// TIA Portal V21 export
// export: Created 2026-08-21T20:18:52.6792221Z, ExportSetting None, DisplayName Totally Integrated Automation Portal, DisplayVersion V21, DisplayName STEP 7 Professional, DisplayVersion V21, DisplayName STEP 7 Safety, DisplayVersion V21, DisplayName Tech WebApplication, DisplayVersion V21, DisplayName WinCC Basic/Comfort/Advanced, DisplayVersion V21, DisplayName WinCC Professional, DisplayVersion V21, DisplayName WinCC Unified, DisplayVersion V21
FUNCTION_BLOCK "ServiceMediumParameterHMI"   // FB1754, SCL
TITLE = ServiceMediumParameterHMI
{ S7_Optimized_Access := 'TRUE' }
AUTHOR : Siemens AG
FAMILY : ServiceControl
VERSION : 4.0
// { "TagName" : "" , "TagDescription" : "" }
// stored: MemoryReserve 100, SetENOAutomatically false
   VAR_INPUT
      Id { ExternalAccessible := 'False'; ExternalVisible := 'False'; ExternalWritable := 'False'} : USInt;   // Service parameter ID
      Setup { ExternalAccessible := 'False'; ExternalVisible := 'False'; ExternalWritable := 'False'} : DB_ANY;   // Setup DB used for the service
      ProcedureCur { ExternalAccessible := 'False'; ExternalVisible := 'False'; ExternalWritable := 'False'} : DWord;   // Current Procedure Number
      ProcedureReq { ExternalAccessible := 'False'; ExternalVisible := 'False'; ExternalWritable := 'False'} : DWord;   // Required Procedure Numbar
   END_VAR
   VAR_IN_OUT
      ConfigurationParameterAnalog : Array[*] of "UDT_MTP_AnaServParam";   // Analog configuration parameter
      ConfigurationParameterDigital : Array[*] of "UDT_MTP_DIntServParam";   // Digital configuration parameter
      ConfigurationParameterBinary : Array[*] of "UDT_MTP_BinServParam";   // Binary configuration parameter
      ConfigurationParameterString : Array[*] of "UDT_MTP_StringServParam";   // String configuration parameter
      ProcedureParameterAnalog : Array[*] of "UDT_MTP_AnaServParam";   // Analog configuration parameter / Analog procedure parameter
      ProcedureParameterDigital : Array[*] of "UDT_MTP_DIntServParam";   // Digital configuration parameter / Digital procedure parameter
      ProcedureParameterBinary : Array[*] of "UDT_MTP_BinServParam";   // Binary configuration parameter / Binary procedure parameter
      ProcedureParameterString : Array[*] of "UDT_MTP_StringServParam";   // String configuration parameter / String procedure parameter
      ProcessValueInAnalog : Array[*] of "UDT_MTP_AnaProcessValueIn";   // Analog process value in
      ProcessValueInDigital : Array[*] of "UDT_MTP_DIntProcessValueIn";   // Digital process value in
      ProcessValueInBinary : Array[*] of "UDT_MTP_BinProcessValueIn";   // Binary process value in
      ProcessValueInString : Array[*] of "UDT_MTP_StringProcessValueIn";   // String process value in
      ProcessValueOutAnalog : Array[*] of "UDT_MTP_AnaProcessValueOut";   // Analog process value out
      ProcessValueOutDigital : Array[*] of "UDT_MTP_DIntProcessValueOut";   // Digital process value out
      ProcessValueOutBinary : Array[*] of "UDT_MTP_BinProcessValueOut";   // Binary process value out
      ProcessValueOutString : Array[*] of "UDT_MTP_StringProcessValueOut";   // String process value out
      ReportValueAnalog : Array[*] of "UDT_MTP_AnaReportValue";   // Analog report value
      ReportValueDigital : Array[*] of "UDT_MTP_DIntReportValue";   // Digital report value
      ReportValueBinary : Array[*] of "UDT_MTP_BinReportValue";   // Binary report value
      ReportValueString : Array[*] of "UDT_MTP_StringReportValue";   // String report value
   END_VAR
   VAR
      statTotalConfigParameters { ExternalAccessible := 'False'; ExternalVisible := 'False'; ExternalWritable := 'False'} : Int;   // Total used configuration parameter
      statTotalProcedureParameters { ExternalAccessible := 'False'; ExternalVisible := 'False'; ExternalWritable := 'False'} : Int;   // Total used procedure parameter
      statTotalProcessInValues { ExternalAccessible := 'False'; ExternalVisible := 'False'; ExternalWritable := 'False'} : Int;   // Total used process in values
      statTotalProcessOutValues { ExternalAccessible := 'False'; ExternalVisible := 'False'; ExternalWritable := 'False'} : Int;   // Total used process Out values
      statTotalReportValues { ExternalAccessible := 'False'; ExternalVisible := 'False'; ExternalWritable := 'False'} : Int;   // Total used Report values
      StatConfigAnalog { ExternalAccessible := 'False'; ExternalVisible := 'False'; ExternalWritable := 'False'} : Array[0..#MAPPED_CONFIG_ANALOG] of "UDT_Service_AnaServParam";   // Writable Config analog parameters
      StatConfigDigital { ExternalAccessible := 'False'; ExternalVisible := 'False'; ExternalWritable := 'False'} : Array[0..#MAPPED_CONFIG_DIGITAL] of "UDT_Service_DintServParam";   // Writable Config digital parameters
      StatConfigBinary { ExternalAccessible := 'False'; ExternalVisible := 'False'; ExternalWritable := 'False'} : Array[0..#MAPPED_CONFIG_BINARY] of "UDT_Service_BinServParam";   // Writable Config binary parameters
      StatConfigString { ExternalAccessible := 'False'; ExternalVisible := 'False'; ExternalWritable := 'False'} : Array[0..#MAPPED_CONFIG_STRING] of "UDT_Service_StringServParam";   // Writable Config string parameters
      StatProcedureAnalog { ExternalAccessible := 'False'; ExternalVisible := 'False'; ExternalWritable := 'False'} : Array[0..#MAPPED_PROCEDURE_ANALOG] of "UDT_Service_AnaServParam";   // Writable Config analog parameters
      StatProcedureDigital { ExternalAccessible := 'False'; ExternalVisible := 'False'; ExternalWritable := 'False'} : Array[0..#MAPPED_PROCEDURE_DIGITAL] of "UDT_Service_DintServParam";   // Writable Config digital parameters
      StatProcedureBinary { ExternalAccessible := 'False'; ExternalVisible := 'False'; ExternalWritable := 'False'} : Array[0..#MAPPED_PROCEDURE_BINARY] of "UDT_Service_BinServParam";   // Writable Config binary parameters
      StatProcedureString { ExternalAccessible := 'False'; ExternalVisible := 'False'; ExternalWritable := 'False'} : Array[0..#MAPPED_PROCEDURE_STRING] of "UDT_Service_StringServParam";   // Writable Config string parameters
      stat16ProceReqIndex { ExternalAccessible := 'False'; ExternalVisible := 'False'; ExternalWritable := 'False'} : Int;   // Requested/Prepared procedure index number
      stat16ProceCurIndex { ExternalAccessible := 'False'; ExternalVisible := 'False'; ExternalWritable := 'False'} : Int;   // current/Running procedure index number
      stat16ProcParaStartIndex { ExternalAccessible := 'False'; ExternalVisible := 'False'; ExternalWritable := 'False'} : Int;   // Procedure parameter start index value
      stat16ProcParaEndIndex { ExternalAccessible := 'False'; ExternalVisible := 'False'; ExternalWritable := 'False'} : Int;   // Procedure parameter end index value
      stat32PrecedureProcessOutMap { ExternalAccessible := 'False'; ExternalVisible := 'False'; ExternalWritable := 'False'} : DWord;   // Procedure assignment information for ProcessOut values
      stat32PrecedureProcessInMap { ExternalAccessible := 'False'; ExternalVisible := 'False'; ExternalWritable := 'False'} : DWord;   // Procedure assignment information for ProcessIn values
      stat32PrecedureReportMap { ExternalAccessible := 'False'; ExternalVisible := 'False'; ExternalWritable := 'False'} : DWord;   // Procedure assignment information for Report values
      ConfigParaType : "UDT_Service_ConfigParaIndexType";   // Index information for the configuration parameter
      ProcedureParaType : "UDT_Service_ProceParaValueIndexType";   // Index information for the procedure parameter
      ProcessInValueType : "UDT_Service_ProceParaValueIndexType";   // Index information for the process in values
      ProcessOutValueType : "UDT_Service_ProceParaValueIndexType";   // Index information for the process out values
      ReportValueType : "UDT_Service_ProceParaValueIndexType";   // Index information for the report values
      ConfigAna : Array[0..#MAPPED_CONFIG_ANALOG] of "UDT_MTP_AnaServParam";   // Configuration analog parameter
      ConfigDint : Array[0..#MAPPED_CONFIG_DIGITAL] of "UDT_MTP_DIntServParam";   // Configuration digital parameter
      ConfigBin : Array[0..#MAPPED_CONFIG_BINARY] of "UDT_MTP_BinServParam";   // Configuration binary parameter
      ConfigString : Array[0..#MAPPED_CONFIG_STRING] of "UDT_MTP_StringServParam";   // Configuration string parameter
      ProcedureAna : Array[0..#MAPPED_PROCEDURE_ANALOG] of "UDT_MTP_AnaServParam";   // Procedure analog parameter
      ProcedureDint : Array[0..#MAPPED_PROCEDURE_DIGITAL] of "UDT_MTP_DIntServParam";   // Procedure digital parameter
      ProcedureBin : Array[0..#MAPPED_PROCEDURE_BINARY] of "UDT_MTP_BinServParam";   // Procedure binary parameter
      ProcedureString : Array[0..#MAPPED_PROCEDURE_STRING] of "UDT_MTP_StringServParam";   // Procedure string parameter
      ProcessInAna : Array[0..#MAPPED_PROCESS_IN_ANALOG] of "UDT_MTP_AnaProcessValueIn";   // Process In analog values
      ProcessInDint : Array[0..#MAPPED_PROCESS_IN_DIGITAL] of "UDT_MTP_DIntProcessValueIn";   // Process In digital values
      ProcessInBin : Array[0..#MAPPED_PROCESS_IN_BINARY] of "UDT_MTP_BinProcessValueIn";   // Process In binary values
      ProcessInString : Array[0..#MAPPED_PROCESS_IN_STRING] of "UDT_MTP_StringProcessValueIn";   // Process In string values
      ProcessOutAna : Array[0..#MAPPED_PROCESS_OUT_ANALOG] of "UDT_MTP_AnaProcessValueOut";   // Process Out analog values
      ProcessOutDint : Array[0..#MAPPED_PROCESS_OUT_DIGITAL] of "UDT_MTP_DIntProcessValueOut";   // Process Out digital values
      ProcessOutBin : Array[0..#MAPPED_PROCESS_OUT_BINARY] of "UDT_MTP_BinProcessValueOut";   // Process Out binary values
      ProcessOutString : Array[0..#MAPPED_PROCESS_OUT_STRING] of "UDT_MTP_StringProcessValueOut";   // Process Out string values
      ReportAna : Array[0..#MAPPED_REPORT_ANALOG] of "UDT_MTP_AnaReportValue";   // Report analog values
      ReportDint : Array[0..#MAPPED_REPORT_DIGITAL] of "UDT_MTP_DIntReportValue";   // Report digital values
      ReportBin : Array[0..#MAPPED_REPORT_BINARY] of "UDT_MTP_BinReportValue";   // Report binary values
      ReportString : Array[0..#MAPPED_REPORT_STRING] of "UDT_MTP_StringReportValue";   // Report string values
      statInternalCurProcParameter { ExternalAccessible := 'False'; ExternalVisible := 'False'; ExternalWritable := 'False'} : Array[#PROCEDURE_PARAMETER_MIN..#PROCEDURE_PARAMETER_MAX] of "UDT_Service_Parameter";   // Internal Procedure Parameter
      statLasProcedureCur { ExternalAccessible := 'False'; ExternalVisible := 'False'; ExternalWritable := 'False'} : DWord;   // Last current procedure
      statLasProcedureReq { ExternalAccessible := 'False'; ExternalVisible := 'False'; ExternalWritable := 'False'} : DWord;   // Last Prepared procedure
      statLastReqProcedSelected { ExternalAccessible := 'False'; ExternalVisible := 'False'; ExternalWritable := 'False'} : Bool;   // Last Prepared procedure
      StatLastProceselReport { ExternalAccessible := 'False'; ExternalVisible := 'False'; ExternalWritable := 'False'} : Bool;   // Last procedure page selection in Report values FP
      StatLastProceselProcessOut { ExternalAccessible := 'False'; ExternalVisible := 'False'; ExternalWritable := 'False'} : Bool;   // Last procedure page selection in ProcessOut values FP
      StatLastProceselProcessIn { ExternalAccessible := 'False'; ExternalVisible := 'False'; ExternalWritable := 'False'} : Bool;   // Last procedure page selection in ProcessIn values FP
   END_VAR
   VAR_TEMP
      temp32TempDword1 : DWord;   // Dummy for work
      temp16IndexOfDefinition : Int;   // Index of Definition array / Internal counter variable
      temp16ParameterCMAddress : Int;   // Control module address of parameter
      temp16ParameterType : Int;   // Type of Parameter
      temp16IndexMTP : Int;   // Index of MTP array / Index fo value
      temp16IndexIO : Int;   // Index of IO array / Index fo value
      tempUsed : Array[#NUMBER_OF_CONTROLMODULES_IN_DW_MIN..#NUMBER_OF_CONTROLMODULES_IN_DW] of DWord;   // Array for input value used
      temp16TempInt1 : Int;   // Dummy for work
      temp16TempInt2 : Int;   // Dummy for work
      temp16i : Int;   // Internal counter variable
      temp16Index : Int;   // Index of value / Index fo value
      tempVariant : Variant;   // Internal work variable of type Variant
      temp16ReturnValue : Int;   // Internal work variable for Return Value
      tempSetup : "UDT_Service_ControlBlockMedium";   // Content of DB "ServiceControlBlockMediumSetup"
      tempProcStartIndex : Int;   // Procedure start index
      tempProcEndIndex : Int;   // Procedure end index
      temp16InitIndex : Int;   // Variable is used to initialize the Digital & String para index
      tempProcStartingStartIndex : Int;   // Procedure start index for Starting state
      tempProcStartingEndIndex : Int;   // Procedure end index for Starting state
      tempProcRunningStartIndex : Int;   // Procedure start index for Running state
      tempProcRunningEndIndex : Int;   // Procedure end index for Running state
      tempProcHoldingStartIndex : Int;   // Procedure start index for Holding state
      tempProcHoldingEndIndex : Int;   // Procedure end index for Holding state
      tempProcUnHoldingStartIndex : Int;   // Procedure start index for UnHolding state
      tempProcUnHoldingEndIndex : Int;   // Procedure end index for UnHolding state
      tempProcUnPausingStartIndex : Int;   // Procedure start index for Pausing state
      tempProcUnPausingEndIndex : Int;   // Procedure end index for Pausing state
      tempProcResumingStartIndex : Int;   // Procedure start index for Resuming state
      tempProcResumingEndIndex : Int;   // Procedure end index for Resuming state
      tempProcCompletingStartIndex : Int;   // Procedure start index for Completing state
      tempProcCompletingEndIndex : Int;   // Procedure end index for Completing state
      tempProcStoppingStartIndex : Int;   // Procedure start index for Stopping state
      tempProcStoppingEndIndex : Int;   // Procedure end index for Stopping state
      tempProcAbortingStartIndex : Int;   // Procedure start index for Aborting state
      tempProcAbortingEndIndex : Int;   // Procedure end index for Aborting state
      tempProcResettingStartIndex : Int;   // Procedure start index for Resetting state
      tempProcResettingEndIndex : Int;   // Procedure end index for Resetting state
      temp16IndexOfDefinitionProcessOut : Int;   // Index of Definition array / Internal counter variable
      temp16IndexOfDefinitionProcessIn : Int;   // Index of Definition array / Internal counter variable
      temp16IndexOfDefinitionReport : Int;   // Index of Definition array / Internal counter variable
      temp16IndexAnalog : Int;   // Pointer for the used analog parameter
      temp16IndexDigital : Int;   // Pointer for the used digital parameter
      temp16IndexBinary : Int;   // Pointer for the used binary parameter
      temp16IndexString : Int;   // Pointer for the used string parameter
      temp16ReturnValueOBNum : Int;   // Internal work variable for Return Value
      tempTopSi : SI_none;   // Start-up information of current OB
      tempStartSi : SI_none;   // Start-up information of last started OB
      temp16ObNo : UInt;   // OB number
      xOB_Start : Bool;   // block is running in start OB
      temp16ReturnStatus : Word;   // Internal work variable for Return Value
      tempDTLCurrentTime : DTL;   // Current time stamp
   END_VAR
   VAR CONSTANT
      CONFIG_PARAMETER_MIN : Int := 0;   // Minimum number of configuration parameters (planned number -1 due to ArrayAddressing)
      CONFIG_PARAMETER_MAX : Int := 31;   // Maximum number of configuration parameters (planned number -1 due to ArrayAddressing)
      CONFIG_PARAMETER_ANALOG_MAX : Int := 31;   // Maximum number of analog configuration parameters (planned number -1 due to ArrayAddressing)
      CONFIG_PARAMETER_DIGITAL_MAX : Int := 7;   // Maximum number of digital configuration parameters (planned number -1 due to ArrayAddressing)
      CONFIG_PARAMETER_BINARY_MAX : Int := 31;   // Maximum number of binary configuration parameters (planned number -1 due to ArrayAddressing)
      CONFIG_PARAMETER_STRING_MAX : Int := 7;   // Maximum number of string configuration parameters (planned number -1 due to ArrayAddressing)
      PROCEDURE_PARAMETER_MIN : Int := 0;   // Minimum number of procedure parameters (planned number -1 due to ArrayAddressing)
      PROCEDURE_PARAMETER_MAX : Int := 31;   // Maximum number of procedure parameters (planned number -1 due to ArrayAddressing)
      PROCEDURE_PARAMETER_ANALOG_MAX : Int := 31;   // Maximum number of analog procedure parameters (planned number -1 due to ArrayAddressing)
      PROCEDURE_PARAMETER_DIGITAL_MAX : Int := 7;   // Maximum number of digital procedure parameters (planned number -1 due to ArrayAddressing)
      PROCEDURE_PARAMETER_BINARY_MAX : Int := 31;   // Maximum number of binary procedure parameters (planned number -1 due to ArrayAddressing)
      PROCEDURE_PARAMETER_STRING_MAX : Int := 7;   // Maximum number of string procedure parameters (planned number -1 due to ArrayAddressing)
      NUMBER_OF_CONTROLMODULES_IN_DW_MIN : Int := 0;   // Number of control modules coded in DWords (planned number -1 due to ArrayAddressing)
      NUMBER_OF_CONTROLMODULES_IN_DW : Int := 0;   // Number of control modules coded in DWords (planned number -1 due to ArrayAddressing)
      NUMBER_OF_CONTROLMODULES_MIN : Int := 0;   // Number of control modules (planned number -1 due to ArrayAddressing)
      NUMBER_OF_CONTROLMODULES : Int := 29;   // Number of control modules (planned number -1 due to ArrayAddressing)
      TYPE_NONE : USInt := 0;   // No parameter
      TYPE_ANALOG : USInt := 1;   // Parameter / value type analog
      TYPE_DIGITAL : USInt := 2;   // Parameter / value type digital
      TYPE_BINARY : USInt := 3;   // Parameter / value type binary
      TYPE_STRING : USInt := 4;   // Parameter type string
      NUMBER_OF_PROCEDURES_MIN : Int := 0;   // Number of operations (planned number -1 due to ArrayAddressing)
      NUMBER_OF_PROCEDURES : Int := 15;   // Number of operations (planned number -1 due to ArrayAddressing)
      PARAMETERINDEX_MIN : Int := 0;   // Minimum number of configuration parameters (planned number -1 due to ArrayAddressing)
      PARAMETERINDEX_MAX : Int := 511;   // Maximum number of configuration parameters (planned number -1 due to ArrayAddressing)
      REPORT_VALUES_MIN : Int := 0;   // Minimum number of report values (planned number -1 due to ArrayAddressing)
      REPORT_VALUES_MAX : Int := 31;   // Maximum number of report values (planned number -1 due to ArrayAddressing)
      REPORT_VALUES_ANALOG_MAX : Int := 31;   // Maximum number of analog report values (planned number -1 due to ArrayAddressing)
      REPORT_VALUES_DIGITAL_MAX : Int := 7;   // Maximum number of digital report values (planned number -1 due to ArrayAddressing)
      REPORT_VALUES_BINARY_MAX : Int := 31;   // Maximum number of binary report values (planned number -1 due to ArrayAddressing)
      REPORT_VALUES_STRING_MAX : Int := 7;   // Maximum number of string report values (planned number -1 due to ArrayAddressing)
      PROCESS_VALUES_IN_MIN : Int := 0;   // Minimum number of process values in (planned number -1 due to ArrayAddressing)
      PROCESS_VALUES_IN_MAX : Int := 31;   // Maximum number of process values in (planned number -1 due to ArrayAddressing)
      PROCESS_VALUES_IN_ANALOG_MAX : Int := 31;   // Maximum number of analog process values in (planned number -1 due to ArrayAddressing)
      PROCESS_VALUES_IN_DIGITAL_MAX : Int := 7;   // Maximum number of digital process values in (planned number -1 due to ArrayAddressing)
      PROCESS_VALUES_IN_BINARY_MAX : Int := 31;   // Maximum number of binary process values in (planned number -1 due to ArrayAddressing)
      PROCESS_VALUES_IN_STRING_MAX : Int := 7;   // Maximum number of string process values in (planned number -1 due to ArrayAddressing)
      PROCESS_VALUES_OUT_MIN : Int := 0;   // Minimum number of process values out (planned number -1 due to ArrayAddressing)
      PROCESS_VALUES_OUT_MAX : Int := 31;   // Maximum number of process values out (planned number -1 due to ArrayAddressing)
      PROCESS_VALUES_OUT_ANALOG_MAX : Int := 31;   // Maximum number of analog process values out (planned number -1 due to ArrayAddressing)
      PROCESS_VALUES_OUT_DIGITAL_MAX : Int := 7;   // Maximum number of digital process values out (planned number -1 due to ArrayAddressing)
      PROCESS_VALUES_OUT_BINARY_MAX : Int := 31;   // Maximum number of binary process values out (planned number -1 due to ArrayAddressing)
      PROCESS_VALUES_OUT_STRING_MAX : Int := 7;   // Maximum number of string process values out (planned number -1 due to ArrayAddressing)
      MAPPED_CONFIG_ANALOG : Int := 0;   // Mapped configuration analog parameter count
      MAPPED_CONFIG_DIGITAL : Int := 0;   // Mapped configuration digital parameter count
      MAPPED_CONFIG_BINARY : Int := 1;   // Mapped configuration binary parameter count
      MAPPED_CONFIG_STRING : Int := 0;   // Mapped configuration string parameter count
      MAPPED_PROCEDURE_ANALOG : Int := 2;   // Mapped procedure analog parameter count
      MAPPED_PROCEDURE_DIGITAL : Int := 0;   // Mapped procedure digital parameter count
      MAPPED_PROCEDURE_BINARY : Int := 0;   // Mapped procedure binary parameter count
      MAPPED_PROCEDURE_STRING : Int := 0;   // Mapped procedure string parameter count
      MAPPED_PROCESS_IN_ANALOG : Int := 1;   // Mapped process In analog values count
      MAPPED_PROCESS_IN_DIGITAL : Int := 0;   // Mapped process In Digital values count
      MAPPED_PROCESS_IN_BINARY : Int := 1;   // Mapped process In Binary values count
      MAPPED_PROCESS_IN_STRING : Int := 0;   // Mapped process In String values count
      MAPPED_PROCESS_OUT_ANALOG : Int := 1;   // Mapped process Out analog values count
      MAPPED_PROCESS_OUT_DIGITAL : Int := 0;   // Mapped process Out digital values count
      MAPPED_PROCESS_OUT_BINARY : Int := 0;   // Mapped process Out binary values count
      MAPPED_PROCESS_OUT_STRING : Int := 0;   // Mapped process Out string values count
      MAPPED_REPORT_ANALOG : Int := 1;   // Mapped report analog values count
      MAPPED_REPORT_DIGITAL : Int := 0;   // Mapped report digital values count
      MAPPED_REPORT_BINARY : Int := 0;   // Mapped report binary values count
      MAPPED_REPORT_STRING : Int := 0;   // Mapped report string values count
   END_VAR
BEGIN
       REGION Copyright, Change Log
   (*-----------------------------------------------------------------------------------------------------------------------------
       SIEMENS AG
       © Copyright 2021. All Rights Reserved.
       ---------------------------------------------------------------------------------------------------------------------------
       Limitation of liability
       This software was developed with largest care. However, the author can not
       guarantee, that the software runs under each version of SIMATIC Manager on
       each computer flawlessly. There is no warranty for the software, to the extent
       permitted by applicable law. The copyright holder provides the software
       "as is" without warranty of any kind, either expressed or implied, including,
       but not limited to, the implied warranties of merchantability and fitness
       for a particular purpose. The entire risk as to the quality and performance of
       the software is with you. Should the software prove defective, you assume the
       cost of all necessary servicing, repair or correction. In no event unless
       required by applicable law will the copyright holder be liable to you for
       damages, including any general, special, incidental or consequential damages
       arising out of the use or inability to use the software (including but not
       limited to loss of data or data being rendered inaccurate or losses sustained
       by you or third parties or a failure of the software to operate with any
       other programs), even if such holder or other party has been advised of the
       possibility of such damages. Permission to use or copy this software for any
       purpose is hereby granted without fee, provided the above notices are retained
       on all copies. Permission to modify the code and to distribute modified code
       is granted, provided the above notices are retained, and a notice that the
       code was modified is included with the above copyright notice.
       ---------------------------------------------------------------------------------------------------------------------------
       Functionality provided by this source (short description):
       Function block to handle the Parameters mapped/used in the project from the engineering tool.
       ---------------------------------------------------------------------------------------------------------------------------
       Status: Preliminary,
       Preliminary (experimental)
       Baselined  
       Released
       ---------------------------------------------------------------------------------------------------------------------------
       File name:              ServiceParameter.SCL
       Function block name:    "ServiceParameterFB"
       System :                SIMATIC S7 CPU (1500)
       ---------------------------------------------------------------------------------------------------------------------------
       Restrictions, known limitations: (e.g. only for certain platforms, ...)
       The provided source code is applicable to the CPUs of the S7 1500 series
       ---------------------------------------------------------------------------------------------------------------------------
       Requirements, prerequisites, external resources used: (e.g. hardware,
       technological package, memory needed, other scripts which are included,
       other objects instantiated, other applications (e.g. MS Excel) assumed, ...)
       TIA Version V19
       ---------------------------------------------------------------------------------------------------------------------------
       Change log table (latest change is at the bottom of the list):
        Version  | Date       | Expert in charge        | Changes applied
       ----------|------------|-------------------------|-----------------------------
        00.00.01 | 06.03.2024 | Kumaraguru M            | first implement  
        00.00.11 | 26.03.2024 | Kumaraguru M            | BugFix - 682100 - SPFL Library: When the user creates a procedure without assigning a step in the transit state, and after downloading the file to PLC, PLC goes into STOP mode.  
        03.00.01 | 07.04.2024 | Kumaraguru M            | Feature -676519: Process In value view for Service Control Block 
        03.00.01 | 07.04.2024 | Kumaraguru M            | Feature -676521: Process Out value View for Service Control Block 
        03.00.01 | 07.04.2024 | Kumaraguru M            | Feature -676524: Report Value View for Service Control Block
       ---------------------------------------------------------------------------------------------------------------------------
        27.04.2024 - Changed the FB from Type to Master Copy for Memory and Power Tag Optimization
        08.05.2024 - Change : Bug 702554: SPFL: Service Control Block: In the runtime, when the user has not selected a procedure, then the ProcessIn, Processout, and Report parameters are listed.
        08.05.2024 - Change : Bug 700381: SPFL: SPFL Library: When the user engineers the “ServiceParameterHMI” block icon, the interface tag names are not in uniform.
        12.05.2024 - Change : Bug 702859: SPFL: Service Control Block: In the configuration windows, the parameter values are continuously updated.
       ---------------------------------------------------------------------------------------------------------------------------
       Note:User should not change or modify the logic and interfaces of the Funtion Block.
       ---------------------------------------------------------------------------------------------------------------------------*)
       END_REGION

       REGION Get start information / time information
           #temp16ReturnValueOBNum := RD_SINFO(TOP_SI => #tempTopSi, START_UP_SI => #tempStartSi);
           #temp16ObNo := #tempTopSi.OB_Nr;
           #xOB_Start := false;
           IF (#temp16ObNo = 100) THEN
               #xOB_Start := true;
           END_IF;
           #temp16ReturnStatus := INT_TO_WORD(RD_SYS_T(#tempDTLCurrentTime));

       END_REGION

       REGION Initialization
           IF (#temp16ObNo = 100) THEN
               //Reset Config para index
               #ConfigParaType.IndexAnalog := 16#0;
               #ConfigParaType.IndexDigital := 16#0;
               #ConfigParaType.IndexBinary := 16#0;
               #ConfigParaType.IndexString := 16#0;
               //Reset Procedure para index
               #ProcedureParaType.IndexAnalog := 16#0;
               #ProcedureParaType.NameIndexAnalog := 16#0;
               #ProcedureParaType.IndexDigital := 16#0;
               #ProcedureParaType.NameIndexDigital := 16#0;
               #ProcedureParaType.IndexBinary := 16#0;
               #ProcedureParaType.NameIndexBinary := 16#0;
               #ProcedureParaType.IndexString := 16#0;
               #ProcedureParaType.NameIndexString := 16#0;
               //Reset ProcessIn Value index
               #ProcessInValueType.IndexAnalog := 16#0;
               #ProcessInValueType.NameIndexAnalog := 16#0;
               #ProcessInValueType.IndexDigital := 16#0;
               #ProcessInValueType.NameIndexDigital := 16#0;
               #ProcessInValueType.IndexBinary := 16#0;
               #ProcessInValueType.NameIndexBinary := 16#0;
               #ProcessInValueType.IndexString := 16#0;
               #ProcessInValueType.NameIndexString := 16#0;
               //Reset ProcessOut Value index
               #ProcessOutValueType.IndexAnalog := 16#0;
               #ProcessOutValueType.NameIndexAnalog := 16#0;
               #ProcessOutValueType.IndexDigital := 16#0;
               #ProcessOutValueType.NameIndexDigital := 16#0;
               #ProcessOutValueType.IndexBinary := 16#0;
               #ProcessOutValueType.NameIndexBinary := 16#0;
               #ProcessOutValueType.IndexString := 16#0;
               #ProcessOutValueType.NameIndexString := 16#0;
               //Reset Report Value index
               #ReportValueType.IndexAnalog := 16#0;
               #ReportValueType.NameIndexAnalog := 16#0;
               #ReportValueType.IndexDigital := 16#0;
               #ReportValueType.NameIndexDigital := 16#0;
               #ReportValueType.IndexBinary := 16#0;
               #ReportValueType.NameIndexBinary := 16#0;
               #ReportValueType.IndexString := 16#0;
               #ReportValueType.NameIndexString := 16#0;

           END_IF;
       END_REGION


       REGION Check DB_ANY of Source
           // Get the Setup DB UDT info from the Setup DB 
           #tempVariant := DB_ANY_TO_VARIANT(in := #Setup, err => #temp16ReturnValue);
           // Validate Setup DB for the service control medium block and move to temp variable
           IF (#temp16ReturnValue = 0) THEN
               IF TypeOf(#tempVariant) = UDT_Service_ControlBlockMedium THEN
                   #temp16ReturnValue := MOVE_BLK_VARIANT(SRC := #tempVariant, COUNT := 1, SRC_INDEX := 0, DEST_INDEX := 0, DEST => #tempSetup);
               END_IF;
           END_IF;
       END_REGION

       REGION Configuration parameters
           //Initialize the used variable values
           #temp32TempDword1 := 16#1;
           #temp16IndexAnalog := 16#0;
           //#ConfigParaType.IndexAnalog := 16#0;
           #temp16IndexDigital := 16#0;
           //#ConfigParaType.IndexDigital := 16#0;
           #temp16IndexBinary := 16#0;
           //#ConfigParaType.IndexBinary := 16#0;
           #temp16IndexString := 16#0;
           //#ConfigParaType.IndexString := 16#0;
           //Used/Mapped parameter count with individual parameter type will written from the Tool
           #statTotalConfigParameters := #MAPPED_CONFIG_ANALOG + #MAPPED_CONFIG_DIGITAL + #MAPPED_CONFIG_BINARY + #MAPPED_CONFIG_STRING - 1;//Calculate the total used parameter
           IF ((#statTotalConfigParameters >= 0) AND (#statTotalConfigParameters <= #CONFIG_PARAMETER_MAX))  THEN
               FOR #temp16IndexOfDefinition := #CONFIG_PARAMETER_MIN TO #statTotalConfigParameters BY 1 DO//32 config parameters for Medium block.
                   #temp16ParameterCMAddress := BYTE_TO_INT(#tempSetup.configurationParameterData.definition[#temp16IndexOfDefinition].controlModule);//Get CM details from the setup DB.
                   #temp16ParameterType := #tempSetup.configurationParameterData.definition[#temp16IndexOfDefinition].type;//Get parameter type from the setup DB.
                   #temp16IndexMTP := #tempSetup.configurationParameterData.definition[#temp16IndexOfDefinition].indexMTP;//Get parameter indexMTP(wrapper DB) from the setup DB.
                   #temp16IndexIO := #tempSetup.configurationParameterData.definition[#temp16IndexOfDefinition].indexIO;//Get parameter indexIO(service block output config parameter) from the setup DB.
                   #tempUsed := #tempSetup.configurationParameterData.used;//Get parameter used info from setup DB
                   //Condition TO check CMs AND parameter types are in the range
                   IF (#temp16ParameterCMAddress <> 255) AND (#temp16ParameterCMAddress >= #NUMBER_OF_CONTROLMODULES_MIN) AND (#temp16ParameterCMAddress <= #NUMBER_OF_CONTROLMODULES)
                       AND (#temp16ParameterType >= #TYPE_NONE) AND (#temp16ParameterType <= #TYPE_STRING) THEN
                       #temp16TempInt1 := #temp16ParameterCMAddress / 32;    //DWORD - Adress
                       #temp16TempInt2 := #temp16ParameterCMAddress MOD 32;  //Bit - Adress
                       //If parameter is forced (FRC) --> Parameter is used
                       IF (((#tempUsed[#temp16TempInt1] AND SHL(IN := #temp32TempDword1, N := INT_TO_UINT(#temp16TempInt2))) <> 0) = TRUE) THEN
                           CASE #temp16ParameterType OF
                                   // If Parameter type = 1(Analog)
                               #TYPE_ANALOG:
                                   REGION Analog
                                       //Bit Masking funtionality for calculate the used Analog parameter
                                       #ConfigParaType.IndexAnalog := #ConfigParaType.IndexAnalog OR SHL(IN := #temp32TempDword1, N := INT_TO_UINT(#temp16IndexOfDefinition));
                                       //Condition to check the config analog parameters are within range 
                                       IF ((#temp16IndexIO >= #CONFIG_PARAMETER_MIN) AND (#temp16IndexIO <= #MAPPED_CONFIG_ANALOG)) THEN
                                           //WinCC Parameter View Faceplate logic
                                           #ConfigAna[#temp16IndexAnalog].WQC := #ConfigurationParameterAnalog[#temp16IndexMTP].WQC;
                                           #ConfigAna[#temp16IndexAnalog].ApplyEn := #ConfigurationParameterAnalog[#temp16IndexMTP].ApplyEn;
                                           #ConfigAna[#temp16IndexAnalog].ApplyInt := #ConfigurationParameterAnalog[#temp16IndexMTP].ApplyInt;
                                           #ConfigAna[#temp16IndexAnalog].StateChannel := #ConfigurationParameterAnalog[#temp16IndexMTP].StateChannel;
                                           #ConfigAna[#temp16IndexAnalog].StateOffAut := #ConfigurationParameterAnalog[#temp16IndexMTP].StateOffAut;
                                           #ConfigAna[#temp16IndexAnalog].StateOpAut := #ConfigurationParameterAnalog[#temp16IndexMTP].StateOpAut;
                                           #ConfigAna[#temp16IndexAnalog].StateAutAut := #ConfigurationParameterAnalog[#temp16IndexMTP].StateAutAut;
                                           #ConfigAna[#temp16IndexAnalog].StateOffAct := #ConfigurationParameterAnalog[#temp16IndexMTP].StateOffAct;
                                           #ConfigAna[#temp16IndexAnalog].StateOpAct := #ConfigurationParameterAnalog[#temp16IndexMTP].StateOpAct;
                                           #ConfigAna[#temp16IndexAnalog].StateAutAct := #ConfigurationParameterAnalog[#temp16IndexMTP].StateAutAct;
                                           #ConfigAna[#temp16IndexAnalog].SrcChannel := #ConfigurationParameterAnalog[#temp16IndexMTP].SrcChannel;
                                           #ConfigAna[#temp16IndexAnalog].SrcExtAut := #ConfigurationParameterAnalog[#temp16IndexMTP].SrcExtAut;
                                           #ConfigAna[#temp16IndexAnalog].SrcIntAut := #ConfigurationParameterAnalog[#temp16IndexMTP].SrcIntAut;
                                           #ConfigAna[#temp16IndexAnalog].SrcIntAct := #ConfigurationParameterAnalog[#temp16IndexMTP].SrcIntAct;
                                           #ConfigAna[#temp16IndexAnalog].SrcExtAct := #ConfigurationParameterAnalog[#temp16IndexMTP].SrcExtAct;
                                           #ConfigAna[#temp16IndexAnalog].VInt := #ConfigurationParameterAnalog[#temp16IndexMTP].VInt;
                                           #ConfigAna[#temp16IndexAnalog].VReq := #ConfigurationParameterAnalog[#temp16IndexMTP].VReq;
                                           #ConfigAna[#temp16IndexAnalog].VOut := #ConfigurationParameterAnalog[#temp16IndexMTP].VOut;
                                           #ConfigAna[#temp16IndexAnalog].VFbk := #ConfigurationParameterAnalog[#temp16IndexMTP].VFbk;
                                           #ConfigAna[#temp16IndexAnalog].VSclMin := #ConfigurationParameterAnalog[#temp16IndexMTP].VSclMin;
                                           #ConfigAna[#temp16IndexAnalog].VSclMax := #ConfigurationParameterAnalog[#temp16IndexMTP].VSclMax;
                                           #ConfigAna[#temp16IndexAnalog].VUnit := #ConfigurationParameterAnalog[#temp16IndexMTP].VUnit;
                                           #ConfigAna[#temp16IndexAnalog].VMin := #ConfigurationParameterAnalog[#temp16IndexMTP].VMin;
                                           #ConfigAna[#temp16IndexAnalog].VMax := #ConfigurationParameterAnalog[#temp16IndexMTP].VMax;
                                           //Write values from WinCC
                                           IF #ConfigurationParameterAnalog[#temp16IndexMTP].OSLevel = #StatConfigAnalog[#temp16IndexAnalog].OSLevel THEN
                                               #ConfigurationParameterAnalog[#temp16IndexMTP].OSLevel := #ConfigAna[#temp16IndexAnalog].OSLevel;
                                           ELSE
                                               #ConfigAna[#temp16IndexAnalog].OSLevel := #ConfigurationParameterAnalog[#temp16IndexMTP].OSLevel;
                                           END_IF;
                                           IF #ConfigurationParameterAnalog[#temp16IndexMTP].ApplyExt = #StatConfigAnalog[#temp16IndexAnalog].ApplyExt THEN
                                               #ConfigurationParameterAnalog[#temp16IndexMTP].ApplyExt := #ConfigAna[#temp16IndexAnalog].ApplyExt;
                                           ELSE
                                               #ConfigAna[#temp16IndexAnalog].ApplyExt := #ConfigurationParameterAnalog[#temp16IndexMTP].ApplyExt;
                                           END_IF;
                                           IF #ConfigurationParameterAnalog[#temp16IndexMTP].ApplyOp = #StatConfigAnalog[#temp16IndexAnalog].ApplyOp THEN
                                               #ConfigurationParameterAnalog[#temp16IndexMTP].ApplyOp := #ConfigAna[#temp16IndexAnalog].ApplyOp;
                                           ELSE
                                               #ConfigAna[#temp16IndexAnalog].ApplyOp := #ConfigurationParameterAnalog[#temp16IndexMTP].ApplyOp;
                                           END_IF;
                                           IF #ConfigurationParameterAnalog[#temp16IndexMTP].Sync = #StatConfigAnalog[#temp16IndexAnalog].Sync THEN
                                               #ConfigurationParameterAnalog[#temp16IndexMTP].Sync := #ConfigAna[#temp16IndexAnalog].Sync;
                                           ELSE
                                               #ConfigAna[#temp16IndexAnalog].Sync := #ConfigurationParameterAnalog[#temp16IndexMTP].Sync;
                                           END_IF;
                                           IF #ConfigurationParameterAnalog[#temp16IndexMTP].StateOffOp = #StatConfigAnalog[#temp16IndexAnalog].StateOffOp THEN
                                               #ConfigurationParameterAnalog[#temp16IndexMTP].StateOffOp := #ConfigAna[#temp16IndexAnalog].StateOffOp;
                                           ELSE
                                               #ConfigAna[#temp16IndexAnalog].StateOffOp := #ConfigurationParameterAnalog[#temp16IndexMTP].StateOffOp;
                                           END_IF;
                                           IF #ConfigurationParameterAnalog[#temp16IndexMTP].StateOpOp = #StatConfigAnalog[#temp16IndexAnalog].StateOpOp THEN
                                               #ConfigurationParameterAnalog[#temp16IndexMTP].StateOpOp := #ConfigAna[#temp16IndexAnalog].StateOpOp;
                                           ELSE
                                               #ConfigAna[#temp16IndexAnalog].StateOpOp := #ConfigurationParameterAnalog[#temp16IndexMTP].StateOpOp;
                                           END_IF;
                                           IF #ConfigurationParameterAnalog[#temp16IndexMTP].StateAutOp = #StatConfigAnalog[#temp16IndexAnalog].StateAutOp THEN
                                               #ConfigurationParameterAnalog[#temp16IndexMTP].StateAutOp := #ConfigAna[#temp16IndexAnalog].StateAutOp;
                                           ELSE
                                               #ConfigAna[#temp16IndexAnalog].StateAutOp := #ConfigurationParameterAnalog[#temp16IndexMTP].StateAutOp;
                                           END_IF;
                                           IF #ConfigurationParameterAnalog[#temp16IndexMTP].SrcIntOp = #StatConfigAnalog[#temp16IndexAnalog].SrcIntOp THEN
                                               #ConfigurationParameterAnalog[#temp16IndexMTP].SrcIntOp := #ConfigAna[#temp16IndexAnalog].SrcIntOp;
                                           ELSE
                                               #ConfigAna[#temp16IndexAnalog].SrcIntOp := #ConfigurationParameterAnalog[#temp16IndexMTP].SrcIntOp;
                                           END_IF;
                                           IF #ConfigurationParameterAnalog[#temp16IndexMTP].SrcExtOp = #StatConfigAnalog[#temp16IndexAnalog].SrcExtOp THEN
                                               #ConfigurationParameterAnalog[#temp16IndexMTP].SrcExtOp := #ConfigAna[#temp16IndexAnalog].SrcExtOp;
                                           ELSE
                                               #ConfigAna[#temp16IndexAnalog].SrcExtOp := #ConfigurationParameterAnalog[#temp16IndexMTP].SrcExtOp;
                                           END_IF;
                                           IF #ConfigurationParameterAnalog[#temp16IndexMTP].VExt = #StatConfigAnalog[#temp16IndexAnalog].VExt THEN
                                               #ConfigurationParameterAnalog[#temp16IndexMTP].VExt := #ConfigAna[#temp16IndexAnalog].VExt;
                                           ELSE
                                               #ConfigAna[#temp16IndexAnalog].VExt := #ConfigurationParameterAnalog[#temp16IndexMTP].VExt;
                                           END_IF;
                                           IF #ConfigurationParameterAnalog[#temp16IndexMTP].VOp = #StatConfigAnalog[#temp16IndexAnalog].VOp THEN
                                               #ConfigurationParameterAnalog[#temp16IndexMTP].VOp := #ConfigAna[#temp16IndexAnalog].VOp;
                                           ELSE
                                               #ConfigAna[#temp16IndexAnalog].VOp := #ConfigurationParameterAnalog[#temp16IndexMTP].VOp;
                                           END_IF;

                                           #StatConfigAnalog[#temp16IndexAnalog].OSLevel := #ConfigAna[#temp16IndexAnalog].OSLevel;
                                           #StatConfigAnalog[#temp16IndexAnalog].ApplyExt := #ConfigAna[#temp16IndexAnalog].ApplyExt;
                                           #StatConfigAnalog[#temp16IndexAnalog].ApplyOp := #ConfigAna[#temp16IndexAnalog].ApplyOp;
                                           #StatConfigAnalog[#temp16IndexAnalog].Sync := #ConfigAna[#temp16IndexAnalog].Sync;
                                           #StatConfigAnalog[#temp16IndexAnalog].StateOffOp := #ConfigAna[#temp16IndexAnalog].StateOffOp;
                                           #StatConfigAnalog[#temp16IndexAnalog].StateOpOp := #ConfigAna[#temp16IndexAnalog].StateOpOp;
                                           #StatConfigAnalog[#temp16IndexAnalog].StateAutOp := #ConfigAna[#temp16IndexAnalog].StateAutOp;
                                           #StatConfigAnalog[#temp16IndexAnalog].SrcIntOp := #ConfigAna[#temp16IndexAnalog].SrcIntOp;
                                           #StatConfigAnalog[#temp16IndexAnalog].SrcExtOp := #ConfigAna[#temp16IndexAnalog].SrcExtOp;
                                           #StatConfigAnalog[#temp16IndexAnalog].VExt := #ConfigAna[#temp16IndexAnalog].VExt;
                                           #StatConfigAnalog[#temp16IndexAnalog].VOp := #ConfigAna[#temp16IndexAnalog].VOp;
                                       END_IF;
                                       #temp16IndexAnalog := #temp16IndexAnalog + 1;
                                   END_REGION
                                   // If Parameter type = 2(Digital)
                               #TYPE_DIGITAL:
                                   REGION Digital
                                       //Bit Masking funtionality for calculate the used Digital parameter
                                       #ConfigParaType.IndexDigital := #ConfigParaType.IndexDigital OR SHL(IN := #temp32TempDword1, N := INT_TO_UINT(#temp16IndexOfDefinition));
                                       //Condition to check the config digital parameters are within range 
                                       IF ((#temp16IndexIO >= #CONFIG_PARAMETER_MIN) AND (#temp16IndexIO <= #MAPPED_CONFIG_DIGITAL)) THEN
                                           //WinCC Parameter View Faceplate logic
                                           #ConfigDint[#temp16IndexDigital].WQC := #ConfigurationParameterDigital[#temp16IndexMTP].WQC;
                                           #ConfigDint[#temp16IndexDigital].ApplyEn := #ConfigurationParameterDigital[#temp16IndexMTP].ApplyEn;
                                           #ConfigDint[#temp16IndexDigital].ApplyInt := #ConfigurationParameterDigital[#temp16IndexMTP].ApplyInt;
                                           #ConfigDint[#temp16IndexDigital].StateChannel := #ConfigurationParameterDigital[#temp16IndexMTP].StateChannel;
                                           #ConfigDint[#temp16IndexDigital].StateOffAut := #ConfigurationParameterDigital[#temp16IndexMTP].StateOffAut;
                                           #ConfigDint[#temp16IndexDigital].StateOpAut := #ConfigurationParameterDigital[#temp16IndexMTP].StateOpAut;
                                           #ConfigDint[#temp16IndexDigital].StateAutAut := #ConfigurationParameterDigital[#temp16IndexMTP].StateAutAut;
                                           #ConfigDint[#temp16IndexDigital].StateOffAct := #ConfigurationParameterDigital[#temp16IndexMTP].StateOffAct;
                                           #ConfigDint[#temp16IndexDigital].StateOpAct := #ConfigurationParameterDigital[#temp16IndexMTP].StateOpAct;
                                           #ConfigDint[#temp16IndexDigital].StateAutAct := #ConfigurationParameterDigital[#temp16IndexMTP].StateAutAct;
                                           #ConfigDint[#temp16IndexDigital].SrcChannel := #ConfigurationParameterDigital[#temp16IndexMTP].SrcChannel;
                                           #ConfigDint[#temp16IndexDigital].SrcExtAut := #ConfigurationParameterDigital[#temp16IndexMTP].SrcExtAut;
                                           #ConfigDint[#temp16IndexDigital].SrcIntAut := #ConfigurationParameterDigital[#temp16IndexMTP].SrcIntAut;
                                           #ConfigDint[#temp16IndexDigital].SrcIntAct := #ConfigurationParameterDigital[#temp16IndexMTP].SrcIntAct;
                                           #ConfigDint[#temp16IndexDigital].SrcExtAct := #ConfigurationParameterDigital[#temp16IndexMTP].SrcExtAct;
                                           #ConfigDint[#temp16IndexDigital].VInt := #ConfigurationParameterDigital[#temp16IndexMTP].VInt;
                                           #ConfigDint[#temp16IndexDigital].VReq := #ConfigurationParameterDigital[#temp16IndexMTP].VReq;
                                           #ConfigDint[#temp16IndexDigital].VOut := #ConfigurationParameterDigital[#temp16IndexMTP].VOut;
                                           #ConfigDint[#temp16IndexDigital].VFbk := #ConfigurationParameterDigital[#temp16IndexMTP].VFbk;
                                           #ConfigDint[#temp16IndexDigital].VSclMin := #ConfigurationParameterDigital[#temp16IndexMTP].VSclMin;
                                           #ConfigDint[#temp16IndexDigital].VSclMax := #ConfigurationParameterDigital[#temp16IndexMTP].VSclMax;
                                           #ConfigDint[#temp16IndexDigital].VUnit := #ConfigurationParameterDigital[#temp16IndexMTP].VUnit;
                                           #ConfigDint[#temp16IndexDigital].VMin := #ConfigurationParameterDigital[#temp16IndexMTP].VMin;
                                           #ConfigDint[#temp16IndexDigital].VMax := #ConfigurationParameterDigital[#temp16IndexMTP].VMax;
                                           //Write values from WinCC
                                           IF #ConfigurationParameterDigital[#temp16IndexMTP].OSLevel = #StatConfigDigital[#temp16IndexDigital].OSLevel THEN
                                               #ConfigurationParameterDigital[#temp16IndexMTP].OSLevel := #ConfigDint[#temp16IndexDigital].OSLevel;
                                           ELSE
                                               #ConfigDint[#temp16IndexDigital].OSLevel := #ConfigurationParameterDigital[#temp16IndexMTP].OSLevel;
                                           END_IF;
                                           IF #ConfigurationParameterDigital[#temp16IndexMTP].ApplyExt = #StatConfigDigital[#temp16IndexDigital].ApplyExt THEN
                                               #ConfigurationParameterDigital[#temp16IndexMTP].ApplyExt := #ConfigDint[#temp16IndexDigital].ApplyExt;
                                           ELSE
                                               #ConfigDint[#temp16IndexDigital].ApplyExt := #ConfigurationParameterDigital[#temp16IndexMTP].ApplyExt;
                                           END_IF;
                                           IF #ConfigurationParameterDigital[#temp16IndexMTP].ApplyOp = #StatConfigDigital[#temp16IndexDigital].ApplyOp THEN
                                               #ConfigurationParameterDigital[#temp16IndexMTP].ApplyOp := #ConfigDint[#temp16IndexDigital].ApplyOp;
                                           ELSE
                                               #ConfigDint[#temp16IndexDigital].ApplyOp := #ConfigurationParameterDigital[#temp16IndexMTP].ApplyOp;
                                           END_IF;
                                           IF #ConfigurationParameterDigital[#temp16IndexMTP].Sync = #StatConfigDigital[#temp16IndexDigital].Sync THEN
                                               #ConfigurationParameterDigital[#temp16IndexMTP].Sync := #ConfigDint[#temp16IndexDigital].Sync;
                                           ELSE
                                               #ConfigDint[#temp16IndexDigital].Sync := #ConfigurationParameterDigital[#temp16IndexMTP].Sync;
                                           END_IF;
                                           IF #ConfigurationParameterDigital[#temp16IndexMTP].StateOffOp = #StatConfigDigital[#temp16IndexDigital].StateOffOp THEN
                                               #ConfigurationParameterDigital[#temp16IndexMTP].StateOffOp := #ConfigDint[#temp16IndexDigital].StateOffOp;
                                           ELSE
                                               #ConfigDint[#temp16IndexDigital].StateOffOp := #ConfigurationParameterDigital[#temp16IndexMTP].StateOffOp;
                                           END_IF;
                                           IF #ConfigurationParameterDigital[#temp16IndexMTP].StateOpOp = #StatConfigDigital[#temp16IndexDigital].StateOpOp THEN
                                               #ConfigurationParameterDigital[#temp16IndexMTP].StateOpOp := #ConfigDint[#temp16IndexDigital].StateOpOp;
                                           ELSE
                                               #ConfigDint[#temp16IndexDigital].StateOpOp := #ConfigurationParameterDigital[#temp16IndexMTP].StateOpOp;
                                           END_IF;
                                           IF #ConfigurationParameterDigital[#temp16IndexMTP].StateAutOp = #StatConfigDigital[#temp16IndexDigital].StateAutOp THEN
                                               #ConfigurationParameterDigital[#temp16IndexMTP].StateAutOp := #ConfigDint[#temp16IndexDigital].StateAutOp;
                                           ELSE
                                               #ConfigDint[#temp16IndexDigital].StateAutOp := #ConfigurationParameterDigital[#temp16IndexMTP].StateAutOp;
                                           END_IF;
                                           IF #ConfigurationParameterDigital[#temp16IndexMTP].SrcIntOp = #StatConfigDigital[#temp16IndexDigital].SrcIntOp THEN
                                               #ConfigurationParameterDigital[#temp16IndexMTP].SrcIntOp := #ConfigDint[#temp16IndexDigital].SrcIntOp;
                                           ELSE
                                               #ConfigDint[#temp16IndexDigital].SrcIntOp := #ConfigurationParameterDigital[#temp16IndexMTP].SrcIntOp;
                                           END_IF;
                                           IF #ConfigurationParameterDigital[#temp16IndexMTP].SrcExtOp = #StatConfigDigital[#temp16IndexDigital].SrcExtOp THEN
                                               #ConfigurationParameterDigital[#temp16IndexMTP].SrcExtOp := #ConfigDint[#temp16IndexDigital].SrcExtOp;
                                           ELSE
                                               #ConfigDint[#temp16IndexDigital].SrcExtOp := #ConfigurationParameterDigital[#temp16IndexMTP].SrcExtOp;
                                           END_IF;
                                           IF #ConfigurationParameterDigital[#temp16IndexMTP].VExt = #StatConfigDigital[#temp16IndexDigital].VExt THEN
                                               #ConfigurationParameterDigital[#temp16IndexMTP].VExt := #ConfigDint[#temp16IndexDigital].VExt;
                                           ELSE
                                               #ConfigDint[#temp16IndexDigital].VExt := #ConfigurationParameterDigital[#temp16IndexMTP].VExt;
                                           END_IF;
                                           IF #ConfigurationParameterDigital[#temp16IndexMTP].VOp = #StatConfigDigital[#temp16IndexDigital].VOp THEN
                                               #ConfigurationParameterDigital[#temp16IndexMTP].VOp := #ConfigDint[#temp16IndexDigital].VOp;
                                           ELSE
                                               #ConfigDint[#temp16IndexDigital].VOp := #ConfigurationParameterDigital[#temp16IndexMTP].VOp;
                                           END_IF;

                                           #StatConfigDigital[#temp16IndexDigital].OSLevel := #ConfigDint[#temp16IndexDigital].OSLevel;
                                           #StatConfigDigital[#temp16IndexDigital].ApplyExt := #ConfigDint[#temp16IndexDigital].ApplyExt;
                                           #StatConfigDigital[#temp16IndexDigital].ApplyOp := #ConfigDint[#temp16IndexDigital].ApplyOp;
                                           #StatConfigDigital[#temp16IndexDigital].Sync := #ConfigDint[#temp16IndexDigital].Sync;
                                           #StatConfigDigital[#temp16IndexDigital].StateOffOp := #ConfigDint[#temp16IndexDigital].StateOffOp;
                                           #StatConfigDigital[#temp16IndexDigital].StateOpOp := #ConfigDint[#temp16IndexDigital].StateOpOp;
                                           #StatConfigDigital[#temp16IndexDigital].StateAutOp := #ConfigDint[#temp16IndexDigital].StateAutOp;
                                           #StatConfigDigital[#temp16IndexDigital].SrcIntOp := #ConfigDint[#temp16IndexDigital].SrcIntOp;
                                           #StatConfigDigital[#temp16IndexDigital].SrcExtOp := #ConfigDint[#temp16IndexDigital].SrcExtOp;
                                           #StatConfigDigital[#temp16IndexDigital].VExt := #ConfigDint[#temp16IndexDigital].VExt;
                                           #StatConfigDigital[#temp16IndexDigital].VOp := #ConfigDint[#temp16IndexDigital].VOp;
                                       END_IF;
                                       #temp16IndexDigital := #temp16IndexDigital + 1;
                                   END_REGION
                                   // If Parameter type = 3(Binary)
                               #TYPE_BINARY:
                                   REGION Binary
                                       //Bit Masking funtionality for calculate the used Binary parameter
                                       #ConfigParaType.IndexBinary := #ConfigParaType.IndexBinary OR SHL(IN := #temp32TempDword1, N := INT_TO_UINT(#temp16IndexOfDefinition));
                                       //Condition to check the config binary parameters are within range 
                                       IF ((#temp16IndexIO >= #CONFIG_PARAMETER_MIN) AND (#temp16IndexIO <= #MAPPED_CONFIG_BINARY)) THEN
                                           //WinCC Parameter View Faceplate logic
                                           #ConfigBin[#temp16IndexBinary].WQC := #ConfigurationParameterBinary[#temp16IndexMTP].WQC;
                                           #ConfigBin[#temp16IndexBinary].ApplyEn := #ConfigurationParameterBinary[#temp16IndexMTP].ApplyEn;
                                           #ConfigBin[#temp16IndexBinary].ApplyInt := #ConfigurationParameterBinary[#temp16IndexMTP].ApplyInt;
                                           #ConfigBin[#temp16IndexBinary].StateChannel := #ConfigurationParameterBinary[#temp16IndexMTP].StateChannel;
                                           #ConfigBin[#temp16IndexBinary].StateOffAut := #ConfigurationParameterBinary[#temp16IndexMTP].StateOffAut;
                                           #ConfigBin[#temp16IndexBinary].StateOpAut := #ConfigurationParameterBinary[#temp16IndexMTP].StateOpAut;
                                           #ConfigBin[#temp16IndexBinary].StateAutAut := #ConfigurationParameterBinary[#temp16IndexMTP].StateAutAut;
                                           #ConfigBin[#temp16IndexBinary].StateOffAct := #ConfigurationParameterBinary[#temp16IndexMTP].StateOffAct;
                                           #ConfigBin[#temp16IndexBinary].StateOpAct := #ConfigurationParameterBinary[#temp16IndexMTP].StateOpAct;
                                           #ConfigBin[#temp16IndexBinary].StateAutAct := #ConfigurationParameterBinary[#temp16IndexMTP].StateAutAct;
                                           #ConfigBin[#temp16IndexBinary].SrcChannel := #ConfigurationParameterBinary[#temp16IndexMTP].SrcChannel;
                                           #ConfigBin[#temp16IndexBinary].SrcExtAut := #ConfigurationParameterBinary[#temp16IndexMTP].SrcExtAut;
                                           #ConfigBin[#temp16IndexBinary].SrcIntAut := #ConfigurationParameterBinary[#temp16IndexMTP].SrcIntAut;
                                           #ConfigBin[#temp16IndexBinary].SrcIntAct := #ConfigurationParameterBinary[#temp16IndexMTP].SrcIntAct;
                                           #ConfigBin[#temp16IndexBinary].SrcExtAct := #ConfigurationParameterBinary[#temp16IndexMTP].SrcExtAct;
                                           #ConfigBin[#temp16IndexBinary].VInt := #ConfigurationParameterBinary[#temp16IndexMTP].VInt;
                                           #ConfigBin[#temp16IndexBinary].VReq := #ConfigurationParameterBinary[#temp16IndexMTP].VReq;
                                           #ConfigBin[#temp16IndexBinary].VOut := #ConfigurationParameterBinary[#temp16IndexMTP].VOut;
                                           #ConfigBin[#temp16IndexBinary].VFbk := #ConfigurationParameterBinary[#temp16IndexMTP].VFbk;
                                           #ConfigBin[#temp16IndexBinary].VState0 := #ConfigurationParameterBinary[#temp16IndexMTP].VState0;
                                           #ConfigBin[#temp16IndexBinary].VState1 := #ConfigurationParameterBinary[#temp16IndexMTP].VState1;
                                           //Write values from WinCC
                                           IF #ConfigurationParameterBinary[#temp16IndexMTP].OSLevel = #StatConfigBinary[#temp16IndexBinary].OSLevel THEN
                                               #ConfigurationParameterBinary[#temp16IndexMTP].OSLevel := #ConfigBin[#temp16IndexBinary].OSLevel;
                                           ELSE
                                               #ConfigBin[#temp16IndexBinary].OSLevel := #ConfigurationParameterBinary[#temp16IndexMTP].OSLevel;
                                           END_IF;
                                           IF #ConfigurationParameterBinary[#temp16IndexMTP].ApplyExt = #StatConfigBinary[#temp16IndexBinary].ApplyExt THEN
                                               #ConfigurationParameterBinary[#temp16IndexMTP].ApplyExt := #ConfigBin[#temp16IndexBinary].ApplyExt;
                                           ELSE
                                               #ConfigBin[#temp16IndexBinary].ApplyExt := #ConfigurationParameterBinary[#temp16IndexMTP].ApplyExt;
                                           END_IF;
                                           IF #ConfigurationParameterBinary[#temp16IndexMTP].ApplyOp = #StatConfigBinary[#temp16IndexBinary].ApplyOp THEN
                                               #ConfigurationParameterBinary[#temp16IndexMTP].ApplyOp := #ConfigBin[#temp16IndexBinary].ApplyOp;
                                           ELSE
                                               #ConfigBin[#temp16IndexBinary].ApplyOp := #ConfigurationParameterBinary[#temp16IndexMTP].ApplyOp;
                                           END_IF;
                                           IF #ConfigurationParameterBinary[#temp16IndexMTP].Sync = #StatConfigBinary[#temp16IndexBinary].Sync THEN
                                               #ConfigurationParameterBinary[#temp16IndexMTP].Sync := #ConfigBin[#temp16IndexBinary].Sync;
                                           ELSE
                                               #ConfigBin[#temp16IndexBinary].Sync := #ConfigurationParameterBinary[#temp16IndexMTP].Sync;
                                           END_IF;
                                           IF #ConfigurationParameterBinary[#temp16IndexMTP].StateOffOp = #StatConfigBinary[#temp16IndexBinary].StateOffOp THEN
                                               #ConfigurationParameterBinary[#temp16IndexMTP].StateOffOp := #ConfigBin[#temp16IndexBinary].StateOffOp;
                                           ELSE
                                               #ConfigBin[#temp16IndexBinary].StateOffOp := #ConfigurationParameterBinary[#temp16IndexMTP].StateOffOp;
                                           END_IF;
                                           IF #ConfigurationParameterBinary[#temp16IndexMTP].StateOpOp = #StatConfigBinary[#temp16IndexBinary].StateOpOp THEN
                                               #ConfigurationParameterBinary[#temp16IndexMTP].StateOpOp := #ConfigBin[#temp16IndexBinary].StateOpOp;
                                           ELSE
                                               #ConfigBin[#temp16IndexBinary].StateOpOp := #ConfigurationParameterBinary[#temp16IndexMTP].StateOpOp;
                                           END_IF;
                                           IF #ConfigurationParameterBinary[#temp16IndexMTP].StateAutOp = #StatConfigBinary[#temp16IndexBinary].StateAutOp THEN
                                               #ConfigurationParameterBinary[#temp16IndexMTP].StateAutOp := #ConfigBin[#temp16IndexBinary].StateAutOp;
                                           ELSE
                                               #ConfigBin[#temp16IndexBinary].StateAutOp := #ConfigurationParameterBinary[#temp16IndexMTP].StateAutOp;
                                           END_IF;
                                           IF #ConfigurationParameterBinary[#temp16IndexMTP].SrcIntOp = #StatConfigBinary[#temp16IndexBinary].SrcIntOp THEN
                                               #ConfigurationParameterBinary[#temp16IndexMTP].SrcIntOp := #ConfigBin[#temp16IndexBinary].SrcIntOp;
                                           ELSE
                                               #ConfigBin[#temp16IndexBinary].SrcIntOp := #ConfigurationParameterBinary[#temp16IndexMTP].SrcIntOp;
                                           END_IF;
                                           IF #ConfigurationParameterBinary[#temp16IndexMTP].SrcExtOp = #StatConfigBinary[#temp16IndexBinary].SrcExtOp THEN
                                               #ConfigurationParameterBinary[#temp16IndexMTP].SrcExtOp := #ConfigBin[#temp16IndexBinary].SrcExtOp;
                                           ELSE
                                               #ConfigBin[#temp16IndexBinary].SrcExtOp := #ConfigurationParameterBinary[#temp16IndexMTP].SrcExtOp;
                                           END_IF;
                                           IF #ConfigurationParameterBinary[#temp16IndexMTP].VExt = #StatConfigBinary[#temp16IndexBinary].VExt THEN
                                               #ConfigurationParameterBinary[#temp16IndexMTP].VExt := #ConfigBin[#temp16IndexBinary].VExt;
                                           ELSE
                                               #ConfigBin[#temp16IndexBinary].VExt := #ConfigurationParameterBinary[#temp16IndexMTP].VExt;
                                           END_IF;
                                           IF #ConfigurationParameterBinary[#temp16IndexMTP].VOp = #StatConfigBinary[#temp16IndexBinary].VOp THEN
                                               #ConfigurationParameterBinary[#temp16IndexMTP].VOp := #ConfigBin[#temp16IndexBinary].VOp;
                                           ELSE
                                               #ConfigBin[#temp16IndexBinary].VOp := #ConfigurationParameterBinary[#temp16IndexMTP].VOp;
                                           END_IF;

                                           #StatConfigBinary[#temp16IndexBinary].OSLevel := #ConfigBin[#temp16IndexBinary].OSLevel;
                                           #StatConfigBinary[#temp16IndexBinary].ApplyExt := #ConfigBin[#temp16IndexBinary].ApplyExt;
                                           #StatConfigBinary[#temp16IndexBinary].ApplyOp := #ConfigBin[#temp16IndexBinary].ApplyOp;
                                           #StatConfigBinary[#temp16IndexBinary].Sync := #ConfigBin[#temp16IndexBinary].Sync;
                                           #StatConfigBinary[#temp16IndexBinary].StateOffOp := #ConfigBin[#temp16IndexBinary].StateOffOp;
                                           #StatConfigBinary[#temp16IndexBinary].StateOpOp := #ConfigBin[#temp16IndexBinary].StateOpOp;
                                           #StatConfigBinary[#temp16IndexBinary].StateAutOp := #ConfigBin[#temp16IndexBinary].StateAutOp;
                                           #StatConfigBinary[#temp16IndexBinary].SrcIntOp := #ConfigBin[#temp16IndexBinary].SrcIntOp;
                                           #StatConfigBinary[#temp16IndexBinary].SrcExtOp := #ConfigBin[#temp16IndexBinary].SrcExtOp;
                                           #StatConfigBinary[#temp16IndexBinary].VExt := #ConfigBin[#temp16IndexBinary].VExt;
                                           #StatConfigBinary[#temp16IndexBinary].VOp := #ConfigBin[#temp16IndexBinary].VOp;
                                       END_IF;
                                       #temp16IndexBinary := #temp16IndexBinary + 1;
                                   END_REGION
                                   // If Parameter type = 4(String)
                               #TYPE_STRING:
                                   REGION String
                                       //Bit Masking funtionality for calculate the used String parameter
                                       #ConfigParaType.IndexString := #ConfigParaType.IndexString OR SHL(IN := #temp32TempDword1, N := INT_TO_UINT(#temp16IndexOfDefinition));
                                       //Condition to check the config string parameters are within range 
                                       IF ((#temp16IndexIO >= #CONFIG_PARAMETER_MIN) AND (#temp16IndexIO <= #MAPPED_CONFIG_STRING)) THEN
                                           //WinCC Parameter View Faceplate logic
                                           #ConfigString[#temp16IndexString].WQC := #ConfigurationParameterString[#temp16IndexMTP].WQC;
                                           #ConfigString[#temp16IndexString].ApplyEn := #ConfigurationParameterString[#temp16IndexMTP].ApplyEn;
                                           #ConfigString[#temp16IndexString].ApplyInt := #ConfigurationParameterString[#temp16IndexMTP].ApplyInt;
                                           #ConfigString[#temp16IndexString].StateChannel := #ConfigurationParameterString[#temp16IndexMTP].StateChannel;
                                           #ConfigString[#temp16IndexString].StateOffAut := #ConfigurationParameterString[#temp16IndexMTP].StateOffAut;
                                           #ConfigString[#temp16IndexString].StateOpAut := #ConfigurationParameterString[#temp16IndexMTP].StateOpAut;
                                           #ConfigString[#temp16IndexString].StateAutAut := #ConfigurationParameterString[#temp16IndexMTP].StateAutAut;
                                           #ConfigString[#temp16IndexString].StateOffAct := #ConfigurationParameterString[#temp16IndexMTP].StateOffAct;
                                           #ConfigString[#temp16IndexString].StateOpAct := #ConfigurationParameterString[#temp16IndexMTP].StateOpAct;
                                           #ConfigString[#temp16IndexString].StateAutAct := #ConfigurationParameterString[#temp16IndexMTP].StateAutAct;
                                           #ConfigString[#temp16IndexString].SrcChannel := #ConfigurationParameterString[#temp16IndexMTP].SrcChannel;
                                           #ConfigString[#temp16IndexString].SrcExtAut := #ConfigurationParameterString[#temp16IndexMTP].SrcExtAut;
                                           #ConfigString[#temp16IndexString].SrcIntAut := #ConfigurationParameterString[#temp16IndexMTP].SrcIntAut;
                                           #ConfigString[#temp16IndexString].SrcIntAct := #ConfigurationParameterString[#temp16IndexMTP].SrcIntAct;
                                           #ConfigString[#temp16IndexString].SrcExtAct := #ConfigurationParameterString[#temp16IndexMTP].SrcExtAct;
                                           #ConfigString[#temp16IndexString].VInt := #ConfigurationParameterString[#temp16IndexMTP].VInt;
                                           #ConfigString[#temp16IndexString].VReq := #ConfigurationParameterString[#temp16IndexMTP].VReq;
                                           #ConfigString[#temp16IndexString].VOut := #ConfigurationParameterString[#temp16IndexMTP].VOut;
                                           #ConfigString[#temp16IndexString].VFbk := #ConfigurationParameterString[#temp16IndexMTP].VFbk;
                                           //Write values from WinCC
                                           IF #ConfigurationParameterString[#temp16IndexMTP].OSLevel = #StatConfigString[#temp16IndexString].OSLevel THEN
                                               #ConfigurationParameterString[#temp16IndexMTP].OSLevel := #ConfigString[#temp16IndexString].OSLevel;
                                           ELSE
                                               #ConfigString[#temp16IndexString].OSLevel := #ConfigurationParameterString[#temp16IndexMTP].OSLevel;
                                           END_IF;
                                           IF #ConfigurationParameterString[#temp16IndexMTP].ApplyExt = #StatConfigString[#temp16IndexString].ApplyExt THEN
                                               #ConfigurationParameterString[#temp16IndexMTP].ApplyExt := #ConfigString[#temp16IndexString].ApplyExt;
                                           ELSE
                                               #ConfigString[#temp16IndexString].ApplyExt := #ConfigurationParameterString[#temp16IndexMTP].ApplyExt;
                                           END_IF;
                                           IF #ConfigurationParameterString[#temp16IndexMTP].ApplyOp = #StatConfigString[#temp16IndexString].ApplyOp THEN
                                               #ConfigurationParameterString[#temp16IndexMTP].ApplyOp := #ConfigString[#temp16IndexString].ApplyOp;
                                           ELSE
                                               #ConfigString[#temp16IndexString].ApplyOp := #ConfigurationParameterString[#temp16IndexMTP].ApplyOp;
                                           END_IF;
                                           IF #ConfigurationParameterString[#temp16IndexMTP].Sync = #StatConfigString[#temp16IndexString].Sync THEN
                                               #ConfigurationParameterString[#temp16IndexMTP].Sync := #ConfigString[#temp16IndexString].Sync;
                                           ELSE
                                               #ConfigString[#temp16IndexString].Sync := #ConfigurationParameterString[#temp16IndexMTP].Sync;
                                           END_IF;
                                           IF #ConfigurationParameterString[#temp16IndexMTP].StateOffOp = #StatConfigString[#temp16IndexString].StateOffOp THEN
                                               #ConfigurationParameterString[#temp16IndexMTP].StateOffOp := #ConfigString[#temp16IndexString].StateOffOp;
                                           ELSE
                                               #ConfigString[#temp16IndexString].StateOffOp := #ConfigurationParameterString[#temp16IndexMTP].StateOffOp;
                                           END_IF;
                                           IF #ConfigurationParameterString[#temp16IndexMTP].StateOpOp = #StatConfigString[#temp16IndexString].StateOpOp THEN
                                               #ConfigurationParameterString[#temp16IndexMTP].StateOpOp := #ConfigString[#temp16IndexString].StateOpOp;
                                           ELSE
                                               #ConfigString[#temp16IndexString].StateOpOp := #ConfigurationParameterString[#temp16IndexMTP].StateOpOp;
                                           END_IF;
                                           IF #ConfigurationParameterString[#temp16IndexMTP].StateAutOp = #StatConfigString[#temp16IndexString].StateAutOp THEN
                                               #ConfigurationParameterString[#temp16IndexMTP].StateAutOp := #ConfigString[#temp16IndexString].StateAutOp;
                                           ELSE
                                               #ConfigString[#temp16IndexString].StateAutOp := #ConfigurationParameterString[#temp16IndexMTP].StateAutOp;
                                           END_IF;
                                           IF #ConfigurationParameterString[#temp16IndexMTP].SrcIntOp = #StatConfigString[#temp16IndexString].SrcIntOp THEN
                                               #ConfigurationParameterString[#temp16IndexMTP].SrcIntOp := #ConfigString[#temp16IndexString].SrcIntOp;
                                           ELSE
                                               #ConfigString[#temp16IndexString].SrcIntOp := #ConfigurationParameterString[#temp16IndexMTP].SrcIntOp;
                                           END_IF;
                                           IF #ConfigurationParameterString[#temp16IndexMTP].SrcExtOp = #StatConfigString[#temp16IndexString].SrcExtOp THEN
                                               #ConfigurationParameterString[#temp16IndexMTP].SrcExtOp := #ConfigString[#temp16IndexString].SrcExtOp;
                                           ELSE
                                               #ConfigString[#temp16IndexString].SrcExtOp := #ConfigurationParameterString[#temp16IndexMTP].SrcExtOp;
                                           END_IF;
                                           IF #ConfigurationParameterString[#temp16IndexMTP].VExt = #StatConfigString[#temp16IndexString].VExt THEN
                                               #ConfigurationParameterString[#temp16IndexMTP].VExt := #ConfigString[#temp16IndexString].VExt;
                                           ELSE
                                               #ConfigString[#temp16IndexString].VExt := #ConfigurationParameterString[#temp16IndexMTP].VExt;
                                           END_IF;
                                           IF #ConfigurationParameterString[#temp16IndexMTP].VOp = #StatConfigString[#temp16IndexString].VOp THEN
                                               #ConfigurationParameterString[#temp16IndexMTP].VOp := #ConfigString[#temp16IndexString].VOp;
                                           ELSE
                                               #ConfigString[#temp16IndexString].VOp := #ConfigurationParameterString[#temp16IndexMTP].VOp;
                                           END_IF;

                                           #StatConfigString[#temp16IndexString].OSLevel := #ConfigString[#temp16IndexString].OSLevel;
                                           #StatConfigString[#temp16IndexString].ApplyExt := #ConfigString[#temp16IndexString].ApplyExt;
                                           #StatConfigString[#temp16IndexString].ApplyOp := #ConfigString[#temp16IndexString].ApplyOp;
                                           #StatConfigString[#temp16IndexString].Sync := #ConfigString[#temp16IndexString].Sync;
                                           #StatConfigString[#temp16IndexString].StateOffOp := #ConfigString[#temp16IndexString].StateOffOp;
                                           #StatConfigString[#temp16IndexString].StateOpOp := #ConfigString[#temp16IndexString].StateOpOp;
                                           #StatConfigString[#temp16IndexString].StateAutOp := #ConfigString[#temp16IndexString].StateAutOp;
                                           #StatConfigString[#temp16IndexString].SrcIntOp := #ConfigString[#temp16IndexString].SrcIntOp;
                                           #StatConfigString[#temp16IndexString].SrcExtOp := #ConfigString[#temp16IndexString].SrcExtOp;
                                           #StatConfigString[#temp16IndexString].VExt := #ConfigString[#temp16IndexString].VExt;
                                           #StatConfigString[#temp16IndexString].VOp := #ConfigString[#temp16IndexString].VOp;
                                       END_IF;
                                       #temp16IndexString := #temp16IndexString + 1;
                                   END_REGION
                           END_CASE;
                       END_IF;
                   END_IF;
               END_FOR;
           END_IF;
       END_REGION
      REGION Procedure Parameter
           REGION Get Current/Prepared procedure ID
               //Get Current procedure index number from setup DB
               IF (#ProcedureCur > 0) THEN
                   FOR #temp16i := #NUMBER_OF_PROCEDURES_MIN TO #NUMBER_OF_PROCEDURES BY 1 DO
                       IF #ProcedureCur = #tempSetup.procedure.procedure[#temp16i].Procedure.ProcedureID THEN
                           #stat16ProceCurIndex := #temp16i;
                           EXIT;
                       END_IF;
                   END_FOR;
               END_IF;
               //Get Prepared procedure index number from setup DB
               IF (#ProcedureReq> 0) THEN
                   FOR #temp16i := #NUMBER_OF_PROCEDURES_MIN TO #NUMBER_OF_PROCEDURES BY 1 DO
                       IF #ProcedureReq = #tempSetup.procedure.procedure[#temp16i].Procedure.ProcedureID THEN
                           #stat16ProceReqIndex := #temp16i;
                           EXIT;
                       END_IF;
                   END_FOR;
               END_IF;
           END_REGION
           REGION Get Start and End index details of the Current /Prepared procedure
               //Current/Prepared procedure selection for parameter display in the faceplate
               IF NOT (#ProcedureParaType.ProcedureReqCurInd) THEN
                   //Get current Procedure step order details from Starting State
                   #tempProcStartingStartIndex := #tempSetup.procedure.procedure[#stat16ProceCurIndex].StateTransient.starting.startIndex;
                   #tempProcStartingEndIndex := #tempSetup.procedure.procedure[#stat16ProceCurIndex].StateTransient.starting.endIndex;
                   //Get current Procedure step order details from Running State
                   #tempProcRunningStartIndex := #tempSetup.procedure.procedure[#stat16ProceCurIndex].StateTransient.running.startIndex;
                   #tempProcRunningEndIndex := #tempSetup.procedure.procedure[#stat16ProceCurIndex].StateTransient.running.endIndex;
                   //Get current Procedure step order details from Holding State
                   #tempProcHoldingStartIndex := #tempSetup.procedure.procedure[#stat16ProceCurIndex].StateTransient.holding.startIndex;
                   #tempProcHoldingEndIndex := #tempSetup.procedure.procedure[#stat16ProceCurIndex].StateTransient.holding.endIndex;
                   //Get current Procedure step order details from unholding State
                   #tempProcUnHoldingStartIndex := #tempSetup.procedure.procedure[#stat16ProceCurIndex].StateTransient.unholding.startIndex;
                   #tempProcUnHoldingEndIndex := #tempSetup.procedure.procedure[#stat16ProceCurIndex].StateTransient.unholding.endIndex;
                   //Get current Procedure step order details from pausing State
                   #tempProcUnPausingStartIndex := #tempSetup.procedure.procedure[#stat16ProceCurIndex].StateTransient.pausing.startIndex;
                   #tempProcUnPausingEndIndex := #tempSetup.procedure.procedure[#stat16ProceCurIndex].StateTransient.pausing.endIndex;
                   //Get current Procedure step order details from resuming State
                   #tempProcResumingStartIndex := #tempSetup.procedure.procedure[#stat16ProceCurIndex].StateTransient.resuming.startIndex;
                   #tempProcResumingEndIndex := #tempSetup.procedure.procedure[#stat16ProceCurIndex].StateTransient.resuming.endIndex;
                   //Get current Procedure step order details from completing State
                   #tempProcCompletingStartIndex := #tempSetup.procedure.procedure[#stat16ProceCurIndex].StateTransient.completing.startIndex;
                   #tempProcCompletingEndIndex := #tempSetup.procedure.procedure[#stat16ProceCurIndex].StateTransient.completing.endIndex;
                   //Get current Procedure step order details from stopping State
                   #tempProcStoppingStartIndex := #tempSetup.procedure.procedure[#stat16ProceCurIndex].StateTransient.stopping.startIndex;
                   #tempProcStoppingEndIndex := #tempSetup.procedure.procedure[#stat16ProceCurIndex].StateTransient.stopping.endIndex;
                   //Get current Procedure step order details from aborting State
                   #tempProcAbortingStartIndex := #tempSetup.procedure.procedure[#stat16ProceCurIndex].StateTransient.aborting.startIndex;
                   #tempProcAbortingEndIndex := #tempSetup.procedure.procedure[#stat16ProceCurIndex].StateTransient.aborting.endIndex;
                   //Get current Procedure step order details from resetting State
                   #tempProcResettingStartIndex := #tempSetup.procedure.procedure[#stat16ProceCurIndex].StateTransient.resetting.startIndex;
                   #tempProcResettingEndIndex := #tempSetup.procedure.procedure[#stat16ProceCurIndex].StateTransient.resetting.endIndex;

               ELSIF (#ProcedureParaType.ProcedureReqCurInd) THEN
                   //Get current Procedure step order details from Starting State
                   #tempProcStartingStartIndex := #tempSetup.procedure.procedure[#stat16ProceReqIndex].StateTransient.starting.startIndex;
                   #tempProcStartingEndIndex := #tempSetup.procedure.procedure[#stat16ProceReqIndex].StateTransient.starting.endIndex;
                   //Get current Procedure step order details from Running State
                   #tempProcRunningStartIndex := #tempSetup.procedure.procedure[#stat16ProceReqIndex].StateTransient.running.startIndex;
                   #tempProcRunningEndIndex := #tempSetup.procedure.procedure[#stat16ProceReqIndex].StateTransient.running.endIndex;
                   //Get current Procedure step order details from Holding State
                   #tempProcHoldingStartIndex := #tempSetup.procedure.procedure[#stat16ProceReqIndex].StateTransient.holding.startIndex;
                   #tempProcHoldingEndIndex := #tempSetup.procedure.procedure[#stat16ProceReqIndex].StateTransient.holding.endIndex;
                   //Get current Procedure step order details from unholding State
                   #tempProcUnHoldingStartIndex := #tempSetup.procedure.procedure[#stat16ProceReqIndex].StateTransient.unholding.startIndex;
                   #tempProcUnHoldingEndIndex := #tempSetup.procedure.procedure[#stat16ProceReqIndex].StateTransient.unholding.endIndex;
                   //Get current Procedure step order details from pausing State
                   #tempProcUnPausingStartIndex := #tempSetup.procedure.procedure[#stat16ProceReqIndex].StateTransient.pausing.startIndex;
                   #tempProcUnPausingEndIndex := #tempSetup.procedure.procedure[#stat16ProceReqIndex].StateTransient.pausing.endIndex;
                   //Get current Procedure step order details from resuming State
                   #tempProcResumingStartIndex := #tempSetup.procedure.procedure[#stat16ProceReqIndex].StateTransient.resuming.startIndex;
                   #tempProcResumingEndIndex := #tempSetup.procedure.procedure[#stat16ProceReqIndex].StateTransient.resuming.endIndex;
                   //Get current Procedure step order details from completing State
                   #tempProcCompletingStartIndex := #tempSetup.procedure.procedure[#stat16ProceReqIndex].StateTransient.completing.startIndex;
                   #tempProcCompletingEndIndex := #tempSetup.procedure.procedure[#stat16ProceReqIndex].StateTransient.completing.endIndex;
                   //Get current Procedure step order details from stopping State
                   #tempProcStoppingStartIndex := #tempSetup.procedure.procedure[#stat16ProceReqIndex].StateTransient.stopping.startIndex;
                   #tempProcStoppingEndIndex := #tempSetup.procedure.procedure[#stat16ProceReqIndex].StateTransient.stopping.endIndex;
                   //Get current Procedure step order details from aborting State
                   #tempProcAbortingStartIndex := #tempSetup.procedure.procedure[#stat16ProceReqIndex].StateTransient.aborting.startIndex;
                   #tempProcAbortingEndIndex := #tempSetup.procedure.procedure[#stat16ProceReqIndex].StateTransient.aborting.endIndex;
                   //Get current Procedure step order details from resetting State
                   #tempProcResettingStartIndex := #tempSetup.procedure.procedure[#stat16ProceReqIndex].StateTransient.resetting.startIndex;
                   #tempProcResettingEndIndex := #tempSetup.procedure.procedure[#stat16ProceReqIndex].StateTransient.resetting.endIndex;
               END_IF;

               #tempProcStartIndex := -1;
               #tempProcEndIndex := -1;
               //Get the Start and End index from the States
               IF (#tempProcStartingStartIndex > -1) AND (#tempProcStartingEndIndex > -1) THEN
                   #tempProcStartIndex := #tempProcStartingStartIndex;
                   #tempProcEndIndex := #tempProcStartingEndIndex;
               ELSIF (#tempProcRunningStartIndex > -1) AND (#tempProcRunningEndIndex > -1) THEN
                   #tempProcStartIndex := #tempProcRunningStartIndex;
                   #tempProcEndIndex := #tempProcRunningEndIndex;
               ELSIF (#tempProcHoldingStartIndex > -1) AND (#tempProcHoldingEndIndex > -1) THEN
                   #tempProcStartIndex := #tempProcHoldingStartIndex;
                   #tempProcEndIndex := #tempProcHoldingEndIndex;
               ELSIF (#tempProcUnHoldingStartIndex > -1) AND (#tempProcUnHoldingEndIndex > -1) THEN
                   #tempProcStartIndex := #tempProcUnHoldingStartIndex;
                   #tempProcEndIndex := #tempProcUnHoldingEndIndex;
               ELSIF (#tempProcUnPausingStartIndex > -1) AND (#tempProcUnPausingEndIndex > -1) THEN
                   #tempProcStartIndex := #tempProcUnPausingStartIndex;
                   #tempProcEndIndex := #tempProcUnPausingEndIndex;
               ELSIF (#tempProcResumingStartIndex > -1) AND (#tempProcResumingEndIndex > -1) THEN
                   #tempProcStartIndex := #tempProcResumingStartIndex;
                   #tempProcEndIndex := #tempProcResumingEndIndex;
               ELSIF (#tempProcCompletingStartIndex > -1) AND (#tempProcCompletingEndIndex > -1) THEN
                   #tempProcStartIndex := #tempProcCompletingStartIndex;
                   #tempProcEndIndex := #tempProcCompletingEndIndex;
               ELSIF (#tempProcStoppingStartIndex > -1) AND (#tempProcStoppingEndIndex > -1) THEN
                   #tempProcStartIndex := #tempProcStoppingStartIndex;
                   #tempProcEndIndex := #tempProcStoppingEndIndex;
               ELSIF (#tempProcAbortingStartIndex > -1) AND (#tempProcAbortingEndIndex > -1) THEN
                   #tempProcStartIndex := #tempProcAbortingStartIndex;
                   #tempProcEndIndex := #tempProcAbortingEndIndex;
               ELSIF (#tempProcResettingStartIndex > -1) AND (#tempProcResettingEndIndex > -1) THEN
                   #tempProcStartIndex := #tempProcResettingStartIndex;
                   #tempProcEndIndex := #tempProcResettingEndIndex;
               END_IF;

               //Get Current Procedure step order parameter index details
               IF (#tempProcStartIndex > -1) AND (#tempProcEndIndex > -1) THEN
                   #stat16ProcParaStartIndex := #tempSetup.stepOrder.stepOrder[#tempProcStartIndex].parameter.startIndex;
                   #stat16ProcParaEndIndex := #tempSetup.stepOrder.stepOrder[#tempProcEndIndex].parameter.endIndex;
               END_IF;
           END_REGION


           REGION Get mapped/used procedure parameters and move to the procedure parameter FP variables
               // Condition to check the start and end index values is within the range
               IF ((#stat16ProcParaStartIndex >= #PARAMETERINDEX_MIN) AND (#stat16ProcParaStartIndex <= #PARAMETERINDEX_MAX))
                   AND ((#stat16ProcParaEndIndex >= #PARAMETERINDEX_MIN) AND (#stat16ProcParaEndIndex <= #PARAMETERINDEX_MAX))
                   AND ((#stat16ProcParaEndIndex - #stat16ProcParaStartIndex + #PROCEDURE_PARAMETER_MIN) <= #PROCEDURE_PARAMETER_MAX) THEN

